// TIA Portal V20 export
TYPE "Zylinder_SMC"
   STRUCT
      Wartungsintervall : DInt;
      Fertigmeldung_Zylinder : Bool;
      Aktorzyklen : DInt;
      Auto_Frg_GS : Bool;
      Auto_Frg_AS : Bool;
      Manu_Frg_GS : Bool;
      Manu_Frg_AS : Bool;
      Einr_Frg_GS : Bool;
      Einr_Frg_AS : Bool;
      Init_Frg_GS : Bool;
      Init_Frg_AS : Bool;
      Richt_Frg_GS : Bool;
      Richt_Frg_AS : Bool;
      M_Zylinder_Sensor_AS : Bool;
      M_Eingang_Sensor_GS_Neg : Bool;
   END_STRUCT;
END_TYPE
